{attribute 'enable_dynamic_creation'}
FUNCTION_BLOCK FB_Number EXTENDS FB_AnyValue IMPLEMENTS I_OtlpValue
VAR_OUTPUT
	value: AnyType;
END_VAR

(*
	Releases this value and clears the caller's pointer to it: call it as p^.delete(pSelf:=p).
	pSelf is cleared before the value is freed, so the caller never keeps a dangling pointer.
	A pointer to any other object is refused and left untouched, and nothing is released.
*)
METHOD delete : BOOL
VAR_IN_OUT
	pSelf: POINTER TO FB_AnyValue;
END_VAR
VAR
	_pThis: POINTER TO FB_Number;
	_pSelfAsParam: POINTER TO FB_AnyValue;
END_VAR
_pThis := THIS;
_pSelfAsParam := _pThis;
IF pSelf <> _pSelfAsParam THEN
	RETURN;
END_IF

pSelf := 0;
__DELETE(_pThis);
delete := TRUE;
END_METHOD

PROPERTY eType : E_ValueType
GET
eType := E_ValueType.E_Number;
END_GET
END_PROPERTY

//FB_Exit must be implemented explicitly. If there is an implementation, then the
//method is called before the controller removes the code of the function block instance
//(implicit call). The return value is not evaluated.
METHOD FB_Exit: BOOL
VAR_INPUT
    bInCopyCode: BOOL;  // TRUE: the exit method is called in order to leave the instance which will be copied afterwards (online change).  
END_VAR
THIS^.free();
END_METHOD

//FB_Init is always available implicitly and it is used primarily for initialization.
//The return value is not evaluated. For a specific influence, you can also declare the
//methods explicitly and provide additional code there with the standard initialization
//code. You can evaluate the return value.
METHOD FB_Init: BOOL
VAR_INPUT
    bInitRetains: BOOL; // TRUE: the retain variables are initialized (reset warm / reset cold)
    bInCopyCode: BOOL;  // TRUE: the instance will be copied to the copy code afterward (online change)
	value: AnyType;
END_VAR
(* ValueFactory owns validation and allocation. FB_Number takes ownership of
the copied value and its type metadata only after every allocation succeeds. *)
THIS^.value := value;
END_METHOD

(* deallocates all data owned by the value without deleting the object itself.*)
METHOD free
IF THIS^.value.pValue <> 0 THEN
	__DELETE(THIS^.value.pValue);
END_IF
MEMSET(ADR(THIS^.value), 0, SIZEOF(THIS^.value));
END_METHOD

END_FUNCTION_BLOCK

(* stored: Version 1.1.0.1
   POU FB_Number: Id {c5fb9a17-5d56-41cb-88c0-bdfb63683555}, SpecialFunc None
   Method delete: Id {81626baf-73e9-474d-8fdb-3db32f627943}
   Property eType: Id {5bc99ae1-764d-46dc-ad39-c02b186a1dfd}
   Get Get: Id {7e33065d-f409-44ce-a7b2-721cf13cf094}
   Method FB_Exit: Id {7b92b00a-edbb-42b3-adc5-8a7e65018ece}
   Method FB_Init: Id {d6aad393-9bab-4c5d-928a-ab98d173ed73}
   Method free: Id {befe6018-20a6-42af-8f70-d8bf62cbbf12} *)
